(* IEC 61131-3 sources: JingjiangMoonbox/Application/Application/数据类型/系统参数/其他参数集/Tension_2024, 7 files *)

(* ---- Cached_Array_Pointers.st ---- *)
(*@CES
Name=Cached_Array_Pointers
Type=Gvl
TypeGuid=2db5746d-d284-4425-9f7f-2663a34b0ebc
Guid=43bd4314-ec4c-41de-8fe2-1da090fdbc31
HasDeclaration=True
HasImplementation=False
*)
{DECLARATION}
TYPE Cached_Array_Pointers :
STRUCT
	(*PI控制器*)
		arUk_PI:ARRAY [1..2] OF REAL;(*输入寄存器*)
		arYk_PI: ARRAY [1..2] OF REAL;(*输出寄存器*)
	(*Kalman*)
	(*上一拍的状态误差协方差矩阵Ph和状态矩阵Xh*)
		arPh:ARRAY [1..4,1..4] OF REAL;(*上一个周期的先验状态误差协方差矩阵*)
		arXh: ARRAY [1..4] OF REAL;(*上一个周期估计状态向量Xh指针*)
	(*LQR迭代求解DARE*)
		arX_DARE:ARRAY [1..4,1..4] OF REAL;(*上一个周期已经迭代收敛的值X_Dare*)

	(*LQR最大迭代次数*)
		iMaxIterateCnt_LQR:INT;

	(*MinBeat最大迭代次数*)
		iMaxIterateCnt_MinBeat:INT;

	(*2024.06.08.150458+lreal类型*)
	(*上一拍的状态误差协方差矩阵Ph和状态矩阵Xh*)
		alrPh:ARRAY [1..4,1..4] OF LREAL;(*上一个周期的先验状态误差协方差矩阵*)
		alrXh: ARRAY [1..4] OF LREAL;(*上一个周期估计状态向量Xh指针*)
	(*LQR迭代求解DARE*)
		alrX_DARE:ARRAY [1..4,1..4] OF LREAL;(*上一个周期已经迭代收敛的值X_Dare*)
END_STRUCT
END_TYPE

{IMPLEMENTATION}

(* ---- Initial_Model_Parameters.st ---- *)
(*@CES
Name=Initial_Model_Parameters
Type=Gvl
TypeGuid=2db5746d-d284-4425-9f7f-2663a34b0ebc
Guid=d7326a99-ac75-4fbf-9581-4e08c3dedfbc
HasDeclaration=True
HasImplementation=False
*)
{DECLARATION}
{attribute 'pack_mode' := '1'}
TYPE Initial_Model_Parameters :
(*共24bytes|增加冗余空间*)
(*该结构体中参数需要保持 不能随意修改大小@2024.05.28.082414*)
STRUCT
    R_0: REAL;             (*初始卷半径m*)
    a0_0: REAL;           (*初始a0*)
    b1_0: REAL;	 	(*初始b1*)
    Wn_0: REAL;	(*初始Wn*)
    Beta_0: REAL;	(*初始Beta*)
    l_0: REAL;		(*初始调整系数l*)
(*	abyReserved:ARRAY [1..26] OF BYTE;*)

END_STRUCT
END_TYPE

{IMPLEMENTATION}

(* ---- Invariant_Parameters.st ---- *)
(*@CES
Name=Invariant_Parameters
Type=Gvl
TypeGuid=2db5746d-d284-4425-9f7f-2663a34b0ebc
Guid=a59fa2b6-149e-4947-99eb-438790530e43
HasDeclaration=True
HasImplementation=False
*)
{DECLARATION}
{attribute 'pack_mode' := '1'}
TYPE Invariant_Parameters :
(*共16bytes|增加冗余空间*)
(*该结构体中参数需要保持 不能随意修改大小@2024.05.28.082414*)
STRUCT
    Ts: REAL;		(*采样时间Ts*)
    Range: REAL;    	(*输出最大量程*)
    Theta: REAL;	(*摆臂偏角范围*)
    K_adj: REAL;		(*模型调整增益*)
(*	abyReserved:ARRAY [1..14] OF BYTE;*)
END_STRUCT
END_TYPE

{IMPLEMENTATION}

(* ---- Kalman_Status_Estimation_And_Feedback.st ---- *)
(*@CES
Name=Kalman_Status_Estimation_And_Feedback
Type=Gvl
TypeGuid=2db5746d-d284-4425-9f7f-2663a34b0ebc
Guid=be73da61-1457-470f-a8cd-978fb9564fdc
HasDeclaration=True
HasImplementation=False
*)
{DECLARATION}
TYPE Kalman_Status_Estimation_And_Feedback :
(*共152bytes|增加冗余空间，该结构体中参数需要保持*)
STRUCT
	R_K:REAL;
	Q:ARRAY [1..4,1..4] OF REAL;
	P0:ARRAY [1..4,1..4] OF REAL;
	N_LQR:REAL;
	Kf:ARRAY [1..4] OF REAL;

	(*2024.06.08.150600+lreal类型*)
	alrQ:ARRAY [1..4,1..4] OF LREAL;
	alrP0:ARRAY [1..4,1..4] OF LREAL;
	alrKf:ARRAY [1..4] OF LREAL;
(*	abyReserved:ARRAY [1..8] OF BYTE;*)
END_STRUCT
END_TYPE

{IMPLEMENTATION}

(* ---- Kalman_Status_Estimation_And_Feedback_MinBeat.st ---- *)
(*@CES
Name=Kalman_Status_Estimation_And_Feedback_MinBeat
Type=Gvl
TypeGuid=2db5746d-d284-4425-9f7f-2663a34b0ebc
Guid=878dded7-317a-4582-b4ff-cfa950f880b6
HasDeclaration=True
HasImplementation=False
*)
{DECLARATION}
TYPE Kalman_Status_Estimation_And_Feedback_MinBeat :
(*共150bytes|增加冗余空间，该结构体中参数需要保持*)
STRUCT
	R_K:REAL;
	Q:ARRAY [1..4,1..4] OF REAL;
	P0:ARRAY [1..4,1..4] OF REAL;
	N_MinBeat:INT;
	Kf:ARRAY [1..4] OF REAL;

(*	abyReserved:ARRAY [1..8] OF BYTE;*)
END_STRUCT
END_TYPE

{IMPLEMENTATION}

(* ---- PI_Parameters.st ---- *)
(*@CES
Name=PI_Parameters
Type=Gvl
TypeGuid=2db5746d-d284-4425-9f7f-2663a34b0ebc
Guid=b0e3524c-689e-4728-99f0-2c6c99433dca
HasDeclaration=True
HasImplementation=False
*)
{DECLARATION}
{attribute 'pack_mode' := '1'}
TYPE PI_Parameters :
(*共12bytes|增加冗余空间*)
(*该结构体中参数需要保持 不能随意修改大小@2024.05.28.082414*)
STRUCT
	(*PI控制器参数*)
	(*K(s+a)/(s+b)*)
	K_PI:REAL;(*系统参数K_PI*)
	a:REAL;(*系统参数a*)
	b:REAL;(*系统参数b*)
(*	abyReserved:ARRAY [1..8] OF BYTE;*)
END_STRUCT
END_TYPE

{IMPLEMENTATION}

(* ---- Time_Varying_Parameters.st ---- *)
(*@CES
Name=Time_Varying_Parameters
Type=Gvl
TypeGuid=2db5746d-d284-4425-9f7f-2663a34b0ebc
Guid=84773baf-ceab-4b75-a59b-2e424c093143
HasDeclaration=True
HasImplementation=False
*)
{DECLARATION}
TYPE Time_Varying_Parameters :
STRUCT
    EST_R: REAL;             	(*卷半径m*)
    a0: REAL;           	(*a0*)
    b1: REAL;	 	(*b1*)
    Wn: REAL;		(*Wn*)
    Beta: REAL;		(*Beta*)
    l: REAL;		(*调整系数l*)
END_STRUCT
END_TYPE

{IMPLEMENTATION}
